Fanuc KAREL source: kt00339.KL

-- PROVISIONAL review KL for V1013-1; original PC SHA256 779d7f0b70c64780b60212ef75d0fb72d32795a8d0bc9abaaa3b5ca16e962457
-- Incomplete behavior may be omitted. Consult companion uncertainty JSON. Do not deploy.
PROGRAM KT00339
%NOLOCKGROUP
VAR
  I2 : INTEGER
  OUT : BOOLEAN
-- UNRESOLVED_DECL Y1 type=002018
BEGIN
  -- UNRESOLVED_PC offsets 5-19; opcodes 2E,22,9D,33,B2
  -- UNRESOLVED_PC offsets 24-35; opcodes 2E,23
  -- UNRESOLVED_PC offsets 40-62; opcodes 22,9D,33,B1,21,59,23
  -- UNRESOLVED_PC offsets 67-71; opcodes 7F
END KT00339
